INTERFACE iSwitch

PROPERTY IsPressed : BOOL
GET
END_GET
END_PROPERTY

PROPERTY IsReleased : BOOL
GET
END_GET
END_PROPERTY

PROPERTY PUBLIC OnPressed : BOOL
GET
END_GET
END_PROPERTY

PROPERTY OnReleased : BOOL
GET
END_GET
END_PROPERTY

END_INTERFACE

(* stored: Version 1.1.0.1
   Itf iSwitch: Id {2b8cdf8a-a619-4e44-ba18-5ff28feae6d7}
   Property IsPressed: Id {36296afe-da41-4462-99a5-b93534c8f214}
   Get Get: Id {822fcb25-a8cd-4415-9cc0-7983d4a3aa52}
   Property IsReleased: Id {95d61822-ed53-4db6-92f9-c11fbffe0b6b}
   Get Get: Id {c3e2ac55-5b65-488d-9296-4e0e905233d0}
   Property OnPressed: Id {76e8bbdf-c484-4aa9-82c0-6b7f3dc3327a}
   Get Get: Id {b1befc1a-e193-4b1a-b19b-81d2f9e2197e}
   Property OnReleased: Id {72547f3f-78f0-4e28-87f6-c436549bb588}
   Get Get: Id {b83f7f50-cdcf-4a72-8eba-03891819d814} *)
